FUNCTION_BLOCK CASE_SEQUENCER (* Migrated from IEC 61131-3 ST *)
  (* Standard: 61499-2 *)
  (* Version 1.0, 2026-11-06, st2fb *)
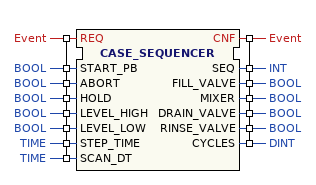
  EVENT_INPUT
    REQ WITH START_PB, ABORT, HOLD, LEVEL_HIGH, LEVEL_LOW, STEP_TIME, SCAN_DT;
  END_EVENT
  EVENT_OUTPUT
    CNF WITH SEQ, FILL_VALVE, MIXER, DRAIN_VALVE, RINSE_VALVE, CYCLES;
  END_EVENT
  VAR_INPUT
    START_PB : BOOL;
    ABORT : BOOL;
    HOLD : BOOL;
    LEVEL_HIGH : BOOL;
    LEVEL_LOW : BOOL;
    STEP_TIME : TIME;
    SCAN_DT : TIME;
  END_VAR
  VAR_OUTPUT
    SEQ : INT;
    FILL_VALVE : BOOL;
    MIXER : BOOL;
    DRAIN_VALVE : BOOL;
    RINSE_VALVE : BOOL;
    CYCLES : DINT;
  END_VAR
  VAR
    TIMING : BOOL := FALSE;
    STEP_TIMER_IN : BOOL := FALSE;
    STEP_TIMER_PT : TIME := T#0s;
    STEP_TIMER_Q : BOOL := FALSE;
    STEP_TIMER_ET : TIME := T#0s;
    STEP_TIMER_STATE : INT := 0;
    STEP_TIMER_PREV_IN : BOOL := FALSE;
    STEP_TIMER_START_TIME : TIME := T#0s;
    ST2FB_NOW : TIME := T#0s;
  END_VAR
  EC_STATES
    START;
    STEP0 : pre, s0 -> CNF;
    W1;
    STEP1 : pre, s1 -> CNF;
    W2;
    STEP2 : pre, s2 -> CNF;
    W3;
    STEP3 : pre, s3 -> CNF;
    W4;
    STEP4 : pre, s4 -> CNF;
    W5;
    STEP5 : pre, s5 -> CNF;
    W6;
    STEP6 : pre, s6 -> CNF;
    W7;
    STEP7 : pre, s7 -> CNF;
    W8;
    STEP8 : pre, s8 -> CNF;
    ABORT_STEP : pre, sabort -> CNF;
  END_STATES
  EC_TRANSITIONS
    START TO ABORT_STEP := REQ[ABORT];
    START TO STEP0 := REQ;
    STEP0 TO W1 := [START_PB];
    STEP0 TO START := 1;
    W1 TO ABORT_STEP := REQ[ABORT];
    W1 TO STEP1 := REQ;
    STEP1 TO W2 := [LEVEL_HIGH];
    STEP1 TO W1 := 1;
    W2 TO ABORT_STEP := REQ[ABORT];
    W2 TO STEP2 := REQ;
    STEP2 TO W3 := [STEP_TIMER_Q];
    STEP2 TO W2 := 1;
    W3 TO ABORT_STEP := REQ[ABORT];
    W3 TO STEP3 := REQ;
    STEP3 TO W4 := [LEVEL_LOW];
    STEP3 TO W3 := 1;
    W4 TO ABORT_STEP := REQ[ABORT];
    W4 TO STEP4 := REQ;
    STEP4 TO W5 := [STEP_TIMER_Q];
    STEP4 TO W4 := 1;
    W5 TO ABORT_STEP := REQ[ABORT];
    W5 TO STEP5 := REQ;
    STEP5 TO W6 := [STEP_TIMER_Q];
    STEP5 TO W5 := 1;
    W6 TO ABORT_STEP := REQ[ABORT];
    W6 TO STEP6 := REQ;
    STEP6 TO W7 := [STEP_TIMER_Q];
    STEP6 TO W6 := 1;
    W7 TO ABORT_STEP := REQ[ABORT];
    W7 TO STEP7 := REQ;
    STEP7 TO START := 1;
    W8 TO ABORT_STEP := REQ[ABORT];
    W8 TO STEP8 := REQ;
    STEP8 TO START := [LEVEL_LOW];
    STEP8 TO W8 := 1;
    ABORT_STEP TO W8 := 1;
  END_TRANSITIONS
  ALGORITHM pre IN ST:
ST2FB_NOW := ST2FB_NOW + SCAN_DT;
IF NOT HOLD THEN
  STEP_TIMER_IN := TIMING;
  STEP_TIMER_PT := STEP_TIME;
  IF (STEP_TIMER_STATE = 0) AND NOT STEP_TIMER_PREV_IN AND STEP_TIMER_IN THEN
    STEP_TIMER_STATE := 1;
    STEP_TIMER_Q := FALSE;
    STEP_TIMER_START_TIME := ST2FB_NOW;
  ELSE
    IF NOT STEP_TIMER_IN THEN
      STEP_TIMER_ET := T#0s;
      STEP_TIMER_Q := FALSE;
      STEP_TIMER_STATE := 0;
    ELSIF STEP_TIMER_STATE = 1 THEN
      IF STEP_TIMER_START_TIME + STEP_TIMER_PT <= ST2FB_NOW THEN
        STEP_TIMER_STATE := 2;
        STEP_TIMER_Q := TRUE;
        STEP_TIMER_ET := STEP_TIMER_PT;
      ELSE
        STEP_TIMER_ET := ST2FB_NOW - STEP_TIMER_START_TIME;
      END_IF;
    END_IF;
  END_IF;
  STEP_TIMER_PREV_IN := STEP_TIMER_IN;
END_IF;
FILL_VALVE := FALSE;
MIXER := FALSE;
DRAIN_VALVE := FALSE;
RINSE_VALVE := FALSE;
  END_ALGORITHM
  ALGORITHM s0 IN ST:
TIMING := FALSE;
IF START_PB THEN
  SEQ := 1;
END_IF;
  END_ALGORITHM
  ALGORITHM s1 IN ST:
FILL_VALVE := TRUE;
IF LEVEL_HIGH THEN
  SEQ := 2;
  TIMING := TRUE;
END_IF;
  END_ALGORITHM
  ALGORITHM s2 IN ST:
MIXER := TRUE;
IF STEP_TIMER_Q THEN
  SEQ := 3;
  TIMING := FALSE;
END_IF;
  END_ALGORITHM
  ALGORITHM s3 IN ST:
DRAIN_VALVE := TRUE;
IF LEVEL_LOW THEN
  SEQ := 4;
END_IF;
  END_ALGORITHM
  ALGORITHM s4 IN ST:
RINSE_VALVE := TRUE;
IF STEP_TIMER_Q THEN
  SEQ := 5;
  TIMING := FALSE;
ELSE
  TIMING := TRUE;
END_IF;
  END_ALGORITHM
  ALGORITHM s5 IN ST:
RINSE_VALVE := TRUE;
IF STEP_TIMER_Q THEN
  SEQ := 6;
  TIMING := FALSE;
ELSE
  TIMING := TRUE;
END_IF;
  END_ALGORITHM
  ALGORITHM s6 IN ST:
RINSE_VALVE := TRUE;
IF STEP_TIMER_Q THEN
  SEQ := 7;
  TIMING := FALSE;
ELSE
  TIMING := TRUE;
END_IF;
  END_ALGORITHM
  ALGORITHM s7 IN ST:
CYCLES := CYCLES + 1;
SEQ := 0;
  END_ALGORITHM
  ALGORITHM s8 IN ST:
TIMING := FALSE;
DRAIN_VALVE := TRUE;
IF LEVEL_LOW AND NOT ABORT THEN
  SEQ := 0;
END_IF;
  END_ALGORITHM
  ALGORITHM sabort IN ST:
SEQ := 8;
TIMING := FALSE;
DRAIN_VALVE := TRUE;
  END_ALGORITHM
END_FUNCTION_BLOCK
